screen "电梯运行监控画面4" 800x600
   Button "按钮_7" at 559,517 size 110x68; TextOff '主画面'
      on Click: ActivateScreen("主画面", 0)
   TextField "文本域_1" at 385,17 size 289x27; Text '-- 4#电梯运行监控'
   TextField "文本域_3" at 114,12 size 263x31; Text '电 梯 监 控 系 统'
   Button "按钮_1" at 678,516 size 106x68; TextOff '退出系统'
      on Click: StopRuntime(0)
   Circle "圆_7" at 199,171 size 31x31
      Appearance <- "输出_4号梯1层按钮指示灯"
   TextField "文本域_9" at 208,175 size 14x19; Text '1'
   Circle "圆_8" at 247,171 size 31x31
      Appearance <- "输出_4号梯2层按钮指示灯"
   TextField "文本域_10" at 256,175 size 14x19; Text '2'
   Circle "圆_9" at 295,171 size 31x31
      Appearance <- "输出_4号梯3层按钮指示灯"
   TextField "文本域_11" at 304,175 size 14x19; Text '3'
   Circle "圆_10" at 199,221 size 31x31
      Appearance <- "输出_4号梯4层按钮指示灯"
   TextField "文本域_12" at 208,225 size 14x19; Text '4'
   Circle "圆_11" at 247,221 size 31x31
      Appearance <- "输出_4号梯5层按钮指示灯"
   TextField "文本域_13" at 256,225 size 14x19; Text '5'
   Circle "圆_12" at 295,221 size 31x31
      Appearance <- "输出_4号梯6层按钮指示灯"
   TextField "文本域_14" at 304,225 size 14x19; Text '6'
   Circle "圆_13" at 199,271 size 31x31
      Appearance <- "输出_4号梯7层按钮指示灯"
   TextField "文本域_15" at 208,275 size 14x19; Text '7'
   Circle "圆_14" at 247,271 size 31x31
      Appearance <- "输出_4号梯8层按钮指示灯"
   TextField "文本域_16" at 256,275 size 14x19; Text '8'
   Circle "圆_15" at 295,271 size 31x31
      Appearance <- "输出_4号梯9层按钮指示灯"
   TextField "文本域_17" at 304,275 size 14x19; Text '9'
   Circle "圆_16" at 248,317 size 31x31
      Appearance <- "输出_4号梯10层按钮指示灯"
   TextField "文本域_18" at 252,322 size 23x19; Text '10'
   TextField "文本域_19" at 368,345 size 61x19; Text '开门'
   TextField "文本域_20" at 457,347 size 53x19; Text '关门'
   TextField "文本域_21" at 528,279 size 95x25; Text '运行方向：'
   TextField "文本域_22" at 529,339 size 94x24; Text '厢门状态：'
   Rectangle "矩形_2" at 178,400 size 599x88
      Visibility <- "输入_4号梯检修信号"
   TextField "文本域_23" at 341,406 size 309x70; Text '4#正常运行'
      Visibility <- "4号梯正常运行"
   GraphicView "图形视图_1" at 609,139 size 124x108; Picture "b_95950E8D4E6480C12C2CE472E64CCEF4[1]"
   Polygon "多边形_3" at 372,298 size 16x33
      Appearance <- "输出_4号梯开门继电器"
   Polygon "多边形_4" at 392,298 size 16x33
      Appearance <- "输出_4号梯开门继电器"
   Polygon "多边形_7" at 459,298 size 16x32
      Appearance <- "输出_4号梯关门继电器"
   Polygon "多边形_8" at 479,298 size 16x32
      Appearance <- "输出_4号梯关门继电器"
   TextField "文本域_24" at 620,293 size 44x19; Text '上行'
      Visibility <- "输出_4号梯上行指示"
   TextField "文本域_25" at 676,291 size 44x19; Text '下行'
      Visibility <- "输出_4号梯下行指示"
   TextField "文本域_27" at 641,352 size 52x19; Text '开启'
      Visibility <- "输出_4号梯开门继电器"
   TextField "文本域_28" at 705,352 size 52x19; Text '关闭'
      Visibility <- "输出_4号梯关门继电器"
   Polygon "多边形_28" at 620,271 size 32x16
      Visibility <- "输出_4号梯上行指示"
   Polygon "多边形_27" at 679,271 size 32x16
      Visibility <- "输出_4号梯下行指示"
   Circle "圆_18" at 652,327 size 21x21
      Visibility <- "输出_4号梯开门继电器"
   Circle "圆_19" at 712,327 size 21x21
      Visibility <- "输出_4号梯关门继电器"
   Button "按钮_2" at 72,133 size 88x45; TextOff 'Text'
      on Click: ActivateScreen("电梯运行监控画面1", 0)
   TextField "文本域_2" at 84,131 size 68x29; Text '1#电梯'
   Button "按钮_3" at 72,189 size 88x45; TextOff 'Text'
      on Click: ActivateScreen("电梯运行监控画面2", 0)
   TextField "文本域_4" at 84,187 size 68x29; Text '2#电梯'
   Button "按钮_4" at 72,247 size 88x45; TextOff 'Text'
      on Click: ActivateScreen("电梯运行监控画面3", 0)
   TextField "文本域_5" at 84,245 size 68x29; Text '3#电梯'
   Button "按钮_5" at 72,305 size 88x45; TextOff 'Text'
      on Click: ActivateScreen("电梯运行监控画面4", 0)
   TextField "文本域_6" at 84,303 size 68x29; Text '4#电梯'
   Button "按钮_6" at 72,363 size 88x45; TextOff 'Text'
      on Click: ActivateScreen("电梯运行监控画面5", 0)
   TextField "文本域_7" at 84,361 size 68x29; Text '5#电梯'
   Button "按钮_8" at 72,421 size 88x45; TextOff 'Text'
      on Click: ActivateScreen("电梯运行监控画面6", 0)
   TextField "文本域_8" at 84,419 size 68x29; Text '6#电梯'
   Rectangle "矩形_193" at 513,169 size 4x18
      Appearance <- "输出_4号梯LEDi"
   Rectangle "矩形_194" at 513,191 size 4x18
      Appearance <- "输出_4号梯LEDj"
   Rectangle "矩形_195" at 526,167 size 18x4
      Appearance <- "输出_4号梯LEDa"
   Rectangle "矩形_196" at 523,171 size 4x18
      Appearance <- "输出_4号梯LEDf"
   Rectangle "矩形_197" at 526,188 size 18x4
      Appearance <- "输出_4号梯LEDg"
   Rectangle "矩形_198" at 523,192 size 4x18
      Appearance <- "输出_4号梯LEDe"
   Rectangle "矩形_199" at 526,210 size 18x4
      Appearance <- "输出_4号梯LEDd"
   Rectangle "矩形_200" at 543,170 size 4x18
      Appearance <- "输出_4号梯LEDb"
   Rectangle "矩形_201" at 543,192 size 4x18
      Appearance <- "输出_4号梯LEDc"
   Rectangle "矩形_72" at 423,156 size 6x34
      Appearance <- "输出_4号梯上行指示"
   Polygon "多边形_5" at 411,152 size 15x17
      Appearance <- "输出_4号梯上行指示"
   Polygon "多边形_6" at 426,152 size 14x17
      Appearance <- "输出_4号梯上行指示"
   Rectangle "矩形_73" at 423,191 size 6x34
      Appearance <- "输出_4号梯下行指示"
   Polygon "多边形_1" at 409,213 size 17x15
      Appearance <- "输出_4号梯下行指示"
   Polygon "多边形_2" at 426,213 size 17x15
      Appearance <- "输出_4号梯下行指示"
   Circle "圆_1" at 21,138 size 35x35
      Appearance <- "1号梯正常运行"
   Circle "圆_2" at 21,194 size 35x35
      Appearance <- "2号梯正常运行"
   Circle "圆_3" at 21,252 size 35x35
      Appearance <- "3号梯正常运行"
   Circle "圆_4" at 21,310 size 35x35
      Appearance <- "4号梯正常运行"
   Circle "圆_5" at 21,368 size 35x35
      Appearance <- "5号梯正常运行"
   Circle "圆_6" at 21,426 size 35x35
      Appearance <- "6号梯正常运行"
   TextField "文本域_33" at 343,403 size 309x70; Text '4#检修故障'
      Visibility <- "输入_4号梯检修信号"
   TextField "文本域_32" at 343,403 size 309x70; Text '4#满载故障'
      Visibility <- "输出_4号梯满载指示"
   Clock "时钟_1" at 664,57 size 101x57
   DateTimeField "日期/时间域_1" at 491,71 size 184x28
   TextField "文本域_26" at 23,498 size 84x47; Text '当前重量'
   IOField "I/O 域_1" at 110,507 size 96x32; FormatPattern s99999
      ProcessValue <- "4号梯载重量"

screen "电梯运行监控画面5" 800x600
   Button "按钮_7" at 559,517 size 110x68; TextOff '主画面'
      on Click: ActivateScreen("主画面", 0)
   TextField "文本域_1" at 385,17 size 284x27; Text '-- 5#电梯运行监控'
   TextField "文本域_3" at 114,12 size 263x31; Text '电 梯 监 控 系 统'
   Button "按钮_1" at 678,516 size 106x68; TextOff '退出系统'
      on Click: StopRuntime(0)
   Circle "圆_7" at 199,171 size 31x31
      Appearance <- "输出_5号梯1层按钮指示灯"
   TextField "文本域_9" at 208,175 size 14x19; Text '1'
   Circle "圆_8" at 247,171 size 31x31
      Appearance <- "输出_5号梯2层按钮指示灯"
   TextField "文本域_10" at 256,175 size 14x19; Text '2'
   Circle "圆_9" at 295,171 size 31x31
      Appearance <- "输出_5号梯3层按钮指示灯"
   TextField "文本域_11" at 304,175 size 14x19; Text '3'
   Circle "圆_10" at 199,221 size 31x31
      Appearance <- "输出_5号梯4层按钮指示灯"
   TextField "文本域_12" at 208,225 size 14x19; Text '4'
   Circle "圆_11" at 247,221 size 31x31
      Appearance <- "输出_5号梯5层按钮指示灯"
   TextField "文本域_13" at 256,225 size 14x19; Text '5'
   Circle "圆_12" at 295,221 size 31x31
      Appearance <- "输出_5号梯6层按钮指示灯"
   TextField "文本域_14" at 304,225 size 14x19; Text '6'
   Circle "圆_13" at 199,271 size 31x31
      Appearance <- "输出_5号梯7层按钮指示灯"
   TextField "文本域_15" at 208,275 size 14x19; Text '7'
   Circle "圆_14" at 247,271 size 31x31
      Appearance <- "输出_5号梯8层按钮指示灯"
   TextField "文本域_16" at 256,275 size 14x19; Text '8'
   Circle "圆_15" at 295,271 size 31x31
      Appearance <- "输出_5号梯9层按钮指示灯"
   TextField "文本域_17" at 304,275 size 14x19; Text '9'
   Circle "圆_16" at 248,317 size 31x31
      Appearance <- "输出_5号梯10层按钮指示灯"
   TextField "文本域_18" at 252,322 size 23x19; Text '10'
   TextField "文本域_19" at 368,345 size 61x19; Text '开门'
   TextField "文本域_20" at 457,347 size 53x19; Text '关门'
   TextField "文本域_21" at 528,279 size 95x25; Text '运行方向：'
   TextField "文本域_22" at 529,339 size 94x24; Text '厢门状态：'
   TextField "文本域_23" at 341,406 size 309x70; Text '5#正常运行'
      Visibility <- "5号梯正常运行"
   GraphicView "图形视图_1" at 609,139 size 124x108; Picture "b_95950E8D4E6480C12C2CE472E64CCEF4[1]"
   Polygon "多边形_3" at 372,298 size 16x33
      Appearance <- "输出_5号梯开门继电器"
   Polygon "多边形_4" at 392,298 size 16x33
      Appearance <- "输出_5号梯开门继电器"
   Polygon "多边形_7" at 459,298 size 16x32
      Appearance <- "输出_5号梯关门继电器"
   Polygon "多边形_8" at 479,298 size 16x32
      Appearance <- "输出_5号梯关门继电器"
   TextField "文本域_24" at 620,289 size 44x19; Text '上行'
      Visibility <- "输出_5号梯上行指示"
   TextField "文本域_25" at 678,287 size 44x19; Text '下行'
      Visibility <- "输出_5号梯下行指示"
   TextField "文本域_27" at 644,348 size 52x19; Text '开启'
      Visibility <- "输出_5号梯开门继电器"
   TextField "文本域_28" at 705,347 size 52x19; Text '关闭'
      Visibility <- "输出_5号梯关门继电器"
   Polygon "多边形_28" at 620,265 size 32x16
      Visibility <- "输出_5号梯上行指示"
   Polygon "多边形_27" at 681,265 size 32x16
      Visibility <- "输出_5号梯下行指示"
   Circle "圆_18" at 652,324 size 21x21
      Visibility <- "输出_5号梯开门继电器"
   Circle "圆_19" at 712,324 size 21x21
      Visibility <- "输出_5号梯关门继电器"
   Button "按钮_2" at 72,133 size 88x45; TextOff 'Text'
      on Click: ActivateScreen("电梯运行监控画面1", 0)
   TextField "文本域_2" at 84,131 size 68x29; Text '1#电梯'
   Button "按钮_3" at 72,189 size 88x45; TextOff 'Text'
      on Click: ActivateScreen("电梯运行监控画面2", 0)
   TextField "文本域_4" at 84,187 size 68x29; Text '2#电梯'
   Button "按钮_4" at 72,247 size 88x45; TextOff 'Text'
      on Click: ActivateScreen("电梯运行监控画面3", 0)
   TextField "文本域_5" at 84,245 size 68x29; Text '3#电梯'
   Button "按钮_5" at 72,305 size 88x45; TextOff 'Text'
      on Click: ActivateScreen("电梯运行监控画面4", 0)
   TextField "文本域_6" at 84,303 size 68x29; Text '4#电梯'
   Button "按钮_6" at 72,363 size 88x45; TextOff 'Text'
      on Click: ActivateScreen("电梯运行监控画面5", 0)
   TextField "文本域_7" at 84,361 size 68x29; Text '5#电梯'
   Button "按钮_8" at 72,421 size 88x45; TextOff 'Text'
      on Click: ActivateScreen("电梯运行监控画面6", 0)
   TextField "文本域_8" at 84,419 size 68x29; Text '6#电梯'
   Rectangle "矩形_193" at 524,172 size 4x18
      Appearance <- "输出_5号梯LEDi"
   Rectangle "矩形_194" at 524,194 size 4x18
      Appearance <- "输出_5号梯LEDj"
   Rectangle "矩形_195" at 537,170 size 18x4
      Appearance <- "输出_5号梯LEDa"
   Rectangle "矩形_196" at 534,174 size 4x18
      Appearance <- "输出_5号梯LEDf"
   Rectangle "矩形_197" at 537,191 size 18x4
      Appearance <- "输出_5号梯LEDg"
   Rectangle "矩形_198" at 534,195 size 4x18
      Appearance <- "输出_5号梯LEDe"
   Rectangle "矩形_199" at 537,213 size 18x4
      Appearance <- "输出_5号梯LEDd"
   Rectangle "矩形_200" at 554,173 size 4x18
      Appearance <- "输出_5号梯LEDb"
   Rectangle "矩形_201" at 554,195 size 4x18
      Appearance <- "输出_5号梯LEDc"
   Rectangle "矩形_72" at 429,160 size 6x34
      Appearance <- "输出_5号梯上行指示"
   Polygon "多边形_5" at 417,156 size 15x17
      Appearance <- "输出_5号梯上行指示"
   Polygon "多边形_6" at 432,156 size 14x17
      Appearance <- "输出_5号梯上行指示"
   Rectangle "矩形_73" at 429,195 size 6x34
      Appearance <- "输出_5号梯下行指示"
   Polygon "多边形_1" at 415,217 size 17x15
      Appearance <- "输出_5号梯下行指示"
   Polygon "多边形_2" at 432,217 size 17x15
      Appearance <- "输出_5号梯下行指示"
   Circle "圆_1" at 21,138 size 35x35
      Appearance <- "1号梯正常运行"
   Circle "圆_2" at 21,194 size 35x35
      Appearance <- "2号梯正常运行"
   Circle "圆_3" at 21,252 size 35x35
      Appearance <- "3号梯正常运行"
   Circle "圆_4" at 21,310 size 35x35
      Appearance <- "4号梯正常运行"
   Circle "圆_5" at 21,368 size 35x35
      Appearance <- "5号梯正常运行"
   Circle "圆_6" at 21,426 size 35x35
      Appearance <- "6号梯正常运行"
   TextField "文本域_33" at 341,408 size 309x70; Text '5#检修故障'
      Visibility <- "输入_5号梯检修信号"
   TextField "文本域_32" at 343,408 size 309x70; Text '5#满载故障'
      Visibility <- "输出_5号梯满载指示"
   Clock "时钟_1" at 664,57 size 101x57
   DateTimeField "日期/时间域_1" at 491,71 size 184x28
   TextField "文本域_26" at 23,498 size 84x47; Text '当前重量'
   IOField "I/O 域_1" at 110,507 size 96x32; FormatPattern s99999
      ProcessValue <- "5号梯载重量"

screen "电梯运行监控画面6" 800x600
   Button "按钮_7" at 559,517 size 110x68; TextOff '主画面'
      on Click: ActivateScreen("主画面", 0)
   TextField "文本域_1" at 385,17 size 295x27; Text '-- 6#电梯运行监控'
   TextField "文本域_3" at 114,12 size 263x31; Text '电 梯 监 控 系 统'
   Button "按钮_1" at 678,516 size 106x68; TextOff '退出系统'
      on Click: StopRuntime(0)
   Circle "圆_7" at 199,171 size 31x31
      Appearance <- "输出_6号梯1层按钮指示灯"
   TextField "文本域_9" at 208,175 size 14x19; Text '1'
   Circle "圆_8" at 247,171 size 31x31
      Appearance <- "输出_6号梯2层按钮指示灯"
   TextField "文本域_10" at 256,175 size 14x19; Text '2'
   Circle "圆_9" at 295,171 size 31x31
      Appearance <- "输出_6号梯3层按钮指示灯"
   TextField "文本域_11" at 304,175 size 14x19; Text '3'
   Circle "圆_10" at 199,221 size 31x31
      Appearance <- "输出_6号梯4层按钮指示灯"
   TextField "文本域_12" at 208,225 size 14x19; Text '4'
   Circle "圆_11" at 247,221 size 31x31
      Appearance <- "输出_6号梯5层按钮指示灯"
   TextField "文本域_13" at 256,225 size 14x19; Text '5'
   Circle "圆_12" at 295,221 size 31x31
      Appearance <- "输出_6号梯6层按钮指示灯"
   TextField "文本域_14" at 304,225 size 14x19; Text '6'
   Circle "圆_13" at 199,271 size 31x31
      Appearance <- "输出_6号梯7层按钮指示灯"
   TextField "文本域_15" at 208,275 size 14x19; Text '7'
   Circle "圆_14" at 247,271 size 31x31
      Appearance <- "输出_6号梯8层按钮指示灯"
   TextField "文本域_16" at 256,275 size 14x19; Text '8'
   Circle "圆_15" at 295,271 size 31x31
      Appearance <- "输出_6号梯9层按钮指示灯"
   TextField "文本域_17" at 304,275 size 14x19; Text '9'
   Circle "圆_16" at 248,317 size 31x31
      Appearance <- "输出_6号梯10层按钮指示灯"
   TextField "文本域_18" at 252,322 size 23x19; Text '10'
   TextField "文本域_19" at 368,345 size 61x19; Text '开门'
   TextField "文本域_20" at 457,347 size 53x19; Text '关门'
   TextField "文本域_21" at 528,280 size 95x25; Text '运行方向：'
   TextField "文本域_22" at 529,340 size 94x24; Text '厢门状态：'
   TextField "文本域_23" at 341,406 size 309x70; Text '6#正常运行'
      Visibility <- "6号梯正常运行"
   GraphicView "图形视图_1" at 609,139 size 124x108; Picture "b_95950E8D4E6480C12C2CE472E64CCEF4[1]"
   Polygon "多边形_3" at 372,298 size 16x33
      Appearance <- "输出_6号梯开门继电器"
   Polygon "多边形_4" at 392,298 size 16x33
      Appearance <- "输出_6号梯开门继电器"
   Polygon "多边形_7" at 459,298 size 16x32
      Appearance <- "输出_6号梯关门继电器"
   Polygon "多边形_8" at 479,298 size 16x32
      Appearance <- "输出_6号梯关门继电器"
   TextField "文本域_24" at 620,288 size 44x19; Text '上行'
      Visibility <- "输出_6号梯上行指示"
   TextField "文本域_25" at 676,286 size 44x19; Text '下行'
      Visibility <- "输出_6号梯下行指示"
   TextField "文本域_27" at 641,349 size 52x19; Text '开启'
      Visibility <- "输出_6号梯开门继电器"
   TextField "文本域_28" at 705,349 size 52x19; Text '关闭'
      Visibility <- "输出_6号梯关门继电器"
   Polygon "多边形_28" at 620,265 size 32x16
      Visibility <- "输出_6号梯上行指示"
   Polygon "多边形_27" at 679,266 size 32x16
      Visibility <- "输出_6号梯下行指示"
   Circle "圆_18" at 652,325 size 21x21
      Visibility <- "输出_6号梯开门继电器"
   Circle "圆_19" at 712,325 size 21x21
      Visibility <- "输出_6号梯关门继电器"
   Button "按钮_2" at 72,133 size 88x45; TextOff 'Text'
      on Click: ActivateScreen("电梯运行监控画面1", 0)
   TextField "文本域_2" at 84,131 size 68x29; Text '1#电梯'
   Button "按钮_3" at 72,189 size 88x45; TextOff 'Text'
      on Click: ActivateScreen("电梯运行监控画面2", 0)
   TextField "文本域_4" at 84,187 size 68x29; Text '2#电梯'
   Button "按钮_4" at 72,247 size 88x45; TextOff 'Text'
      on Click: ActivateScreen("电梯运行监控画面3", 0)
   TextField "文本域_5" at 84,245 size 68x29; Text '3#电梯'
   Button "按钮_5" at 72,305 size 88x45; TextOff 'Text'
      on Click: ActivateScreen("电梯运行监控画面4", 0)
   TextField "文本域_6" at 84,303 size 68x29; Text '4#电梯'
   Button "按钮_6" at 72,363 size 88x45; TextOff 'Text'
      on Click: ActivateScreen("电梯运行监控画面5", 0)
   TextField "文本域_7" at 84,361 size 68x29; Text '5#电梯'
   Button "按钮_8" at 72,421 size 88x45; TextOff 'Text'
      on Click: ActivateScreen("电梯运行监控画面6", 0)
   TextField "文本域_8" at 84,419 size 68x29; Text '6#电梯'
   Rectangle "矩形_193" at 514,170 size 4x18
      Appearance <- "输出_6号梯LEDi"
   Rectangle "矩形_194" at 514,192 size 4x18
      Appearance <- "输出_6号梯LEDj"
   Rectangle "矩形_195" at 527,168 size 18x4
      Appearance <- "输出_6号梯LEDa"
   Rectangle "矩形_196" at 524,172 size 4x18
      Appearance <- "输出_6号梯LEDf"
   Rectangle "矩形_197" at 527,189 size 18x4
      Appearance <- "输出_6号梯LEDg"
   Rectangle "矩形_198" at 524,193 size 4x18
      Appearance <- "输出_6号梯LEDe"
   Rectangle "矩形_199" at 527,211 size 18x4
      Appearance <- "输出_6号梯LEDd"
   Rectangle "矩形_200" at 544,171 size 4x18
      Appearance <- "输出_6号梯LEDb"
   Rectangle "矩形_201" at 544,193 size 4x18
      Appearance <- "输出_6号梯LEDc"
   Rectangle "矩形_72" at 418,157 size 6x34
      Appearance <- "输出_6号梯上行指示"
   Polygon "多边形_5" at 406,153 size 15x17
      Appearance <- "输出_6号梯上行指示"
   Polygon "多边形_6" at 421,153 size 14x17
      Appearance <- "输出_6号梯上行指示"
   Rectangle "矩形_73" at 418,192 size 6x34
      Appearance <- "输出_6号梯下行指示"
   Polygon "多边形_1" at 404,214 size 17x15
      Appearance <- "输出_6号梯下行指示"
   Polygon "多边形_2" at 421,214 size 17x15
      Appearance <- "输出_6号梯下行指示"
   Circle "圆_1" at 21,138 size 35x35
      Appearance <- "1号梯正常运行"
   Circle "圆_2" at 21,194 size 35x35
      Appearance <- "2号梯正常运行"
   Circle "圆_3" at 21,252 size 35x35
      Appearance <- "3号梯正常运行"
   Circle "圆_4" at 21,310 size 35x35
      Appearance <- "4号梯正常运行"
   Circle "圆_5" at 21,368 size 35x35
      Appearance <- "5号梯正常运行"
   Circle "圆_6" at 21,426 size 35x35
      Appearance <- "6号梯正常运行"
   TextField "文本域_33" at 344,408 size 309x70; Text '6#检修故障'
      Visibility <- "输入_6号梯检修信号"
   TextField "文本域_32" at 341,408 size 309x70; Text '6#满载故障'
      Visibility <- "输出_6号梯满载指示"
   Clock "时钟_1" at 664,57 size 101x57
   DateTimeField "日期/时间域_1" at 491,71 size 184x28
   TextField "文本域_26" at 23,498 size 84x47; Text '当前重量'
   IOField "I/O 域_1" at 110,507 size 96x32; FormatPattern s99999
      ProcessValue <- "6号梯载重量"

screen "登录画面" 800x600
   TextField "文本域_1" at 256,120 size 247x74; Text '电梯监控系统'
   Clock "时钟_1" at 690,38 size 101x57
   DateTimeField "日期/时间域_2" at 478,61 size 214x32
   TextField "文本域_2" at 221,217 size 77x21; Text '用户名：'
   TextField "文本域_4" at 229,254 size 69x21; Text '密 码：'
   IOField "I/O 域_1" at 304,259 size 196x25; FormatPattern ????????????????????????????????????????????????????????????????????????????????
      ProcessValue <- "密码"
   IOField "I/O 域_2" at 304,215 size 196x25; FormatPattern ????????????????????????????????????????????????????????????????????????????????
      ProcessValue <- "用户名"
   Button "按钮_3" at 236,319 size 96x32; TextOff '确定'
      on Click: "denglu"(); function_efd93a16("提示信息", 0, 0, -1, -1, 1)
   Button "按钮_4" at 427,319 size 96x32; TextOff '注销'
      on Click: "qingkong"()

screen "设置画面" 800x600
   Button "按钮_7" at 557,516 size 110x66; TextOff '主画面'
      on Click: ActivateScreen("主画面", 0)
   TextField "文本域_1" at 447,16 size 180x27; Text '-- 设置画面'
   TextField "文本域_3" at 130,12 size 263x31; Text '电 梯 监 控 系 统'
   Button "按钮_1" at 677,516 size 106x66; TextOff '退出系统'
      on Click: StopRuntime(0)
   Button "按钮_2" at 275,170 size 243x67; TextOff '初始化楼层设定'
      on Click: ActivateScreen("初始化楼层设定", 0)
   Button "按钮_3" at 274,284 size 243x67; TextOff '用户设置'
      on Click: ActivateScreen("用户设置", 0)
   Clock "时钟_1" at 664,57 size 101x57
   DateTimeField "日期/时间域_1" at 491,71 size 184x28

screen "运行数据记录" 800x600
   Button "按钮_7" at 561,524 size 110x66; TextOff '主画面'
      on Click: ActivateScreen("主画面", 0)
   TextField "文本域_1" at 385,17 size 238x27; Text '-- 电梯状态记录'
   TextField "文本域_3" at 80,12 size 297x31; Text '电 梯 监 控 系 统'
   Button "按钮_1" at 680,524 size 106x66; TextOff '退出系统'
      on Click: StopRuntime(0)
   Clock "时钟_1" at 695,54 size 55x39
   DateTimeField "日期/时间域_1" at 491,59 size 184x28
   RecipeView "配方视图_1" at 156,118 size 400x350; Recipe "配方1"

PopupScreen "提示信息" 500x500
   TextField "文本域_1" at 118,79 size 137x37; Text '提示信息'
   TextField "文本域_3" at 94,146 size 185x19; Text 'Text'
   Button "按钮_1" at 139,194 size 96x32; TextOff '确定'
      on Click: "denglu"()

VB script "denglu"
   '提示：
   ' 1. 使用 <CTRL+SPACE> 或 <CTRL+I> 快捷键打开含所有对象和函数的列表
   ' 2. 使用 HMI Runtime 对象写入代码。
   '  示例：HmiRuntime.Screens("Screen_1")。
   ' 3. 使用 <CTRL+J> 快捷键创建对象引用。
   '从此位置起写入代码：'Please replace all sequences which are enclosed with '_' by your own code.
   
   Dim user,pwd,A
   user=SmartTags("用户名")
   pwd=SmartTags("密码")
   'Please replace all sequences which are enclosed with '_' by your own code.
   If user="admin"And pwd="admin"  Then
   	SmartTags("提示信息")="登录成功"
   	If SmartTags("提示信息")="登录成功"Then
   		A=2
   		acd163fa-ee86-4170-88da-c8d9ec58660c A,0
   	End If
   ElseIf user="" And pwd=""Then
   	SmartTags("提示信息")="错误代码 E0001：用户未登录"
   	If SmartTags("提示信息")="错误代码 E0001：用户未登录"Then
   		A=1
   		acd163fa-ee86-4170-88da-c8d9ec58660c A,0
   	End If
   Else 
   	SmartTags("提示信息")="错误代码 E0002：用户名或密码错误"
   	If SmartTags("提示信息")="错误代码 E0002：用户名或密码错误"Then
   		A=1
   		acd163fa-ee86-4170-88da-c8d9ec58660c A,0
   	End If
   End If

VB script "qingkong"
   '提示：
   ' 1. 使用 <CTRL+SPACE> 或 <CTRL+I> 快捷键打开含所有对象和函数的列表
   ' 2. 使用 HMI Runtime 对象写入代码。
   '  示例：HmiRuntime.Screens("Screen_1")。
   ' 3. 使用 <CTRL+J> 快捷键创建对象引用。
   '从此位置起写入代码：
   SmartTags("用户名")=""
   SmartTags("密码")=""
   SmartTags("提示信息")=""

VB script "tiaozhuan"
   '提示：
   ' 1. 使用 <CTRL+SPACE> 或 <CTRL+I> 快捷键打开含所有对象和函数的列表
   ' 2. 使用 HMI Runtime 对象写入代码。
   '  示例：HmiRuntime.Screens("Screen_1")。
   ' 3. 使用 <CTRL+J> 快捷键创建对象引用。
   '从此位置起写入代码：
   
   'Please replace all sequences which are enclosed with '_' by your own code.
   
   Dim A
   If SmartTags("提示信息")="登录成功"Then
   	A=2
   	acd163fa-ee86-4170-88da-c8d9ec58660c A,0
   End If
   If SmartTags("提示信息")="用户名或密码错误"Then
   	A=1
   	acd163fa-ee86-4170-88da-c8d9ec58660c A,0
   End If

scheduled task "task"
   on Action: function_f41c6f6c("username"); function_e1ab61de("zuhao")
*)